Staubli VAL3: main.pgx

program main()
begin
  close(tCurrentTool)
  pPointRx.config.shoulder = lefty
  pPointRx.config.elbow = epositive
  pPointRx.config.wrist = wpositive
  pPointRx2.config.shoulder = lefty
  pPointRx2.config.elbow = epositive
  pPointRx2.config.wrist = wpositive
  mCurrentSpeed.tvel = 100.00
  mCurrentSpeed.blend = joint
  mCurrentSpeed.reach = 0.010
  mCurrentSpeed.leave = 0.010
  // Program Prog_Name_That_Is_Very_Long_123 start
  // Program generated by VerticalBot Studio for Staubli RX160 on 25/10/2026 12:00:00
  // Using nominal kinematics.
  mCurrentSpeed.tvel = 1000.000
  mCurrentSpeed.reach = 10.000
  mCurrentSpeed.leave = 10.000
  call MoveJoint(10.00000,20.00000,90.00000,30.00000,45.00000,60.00000)
  call MoveLine(1077.300,-56.172,837.243,-146.156,25.288,-102.118)
  mCurrentSpeed.reach = 0.500
  mCurrentSpeed.leave = 0.500
  call MoveLine(1005.190,-118.362,847.372,-147.806,26.655,-97.799)
  delay(0.000)
  delay(1.500)
  popUpMsg("Say "hi" to the operator")
  // A long comment line that exceeds the usual controller limits for comments by far, really
  Output[12]=false
  OUT_A=true
  watch(Input[4]==false,1000.0)
  watch(IN_B==true)
  //call prog:Program_With_A_Long_Name_ABCDEFGHIJ()
  call MoveLine(1077.300,-56.172,837.243,-146.156,25.288,-102.118)
  mCurrentSpeed.reach = -1.000
  mCurrentSpeed.leave = -1.000
  call MoveJoint(10.00000,20.00000,90.00000,30.00000,45.00000,60.00000)

  waitEndMove()
  // Program Prog_Name_That_Is_Very_Long_123 end

end
